Fanuc KAREL source: KO00100.KL

PROGRAM KO00100
%NOLOCKGROUP
VAR
  A: INTEGER
  B: REAL
  OUT: REAL
BEGIN
  A = 1
  B = 2
  OUT = ATAN2(A, B)
END KO00100
